(* IEC 61131-3 sources: LASAL/Drive, 5 files *)

(* ---- _DriveAxis1.st ---- *)
FUNCTION GLOBAL TAB DRIVETAB__DRIVEAXIS1
	1$UDINT, TO_UDINT(OFF(L1)-OFF(L0)),L0:
G01:	1$USINT,'U''C''3'' ',
	2$USINT,' '' '' '' ',
	3$USINT,'3''4''V'' ',
	4$USINT,870$DINT,
	5$USINT,3100$DINT,
	6$USINT,12000$DINT,
	7$USINT,2$DINT,
	8$USINT,30$DINT,
	9$USINT,1950$DINT,
	10$USINT,9400$DINT,
	11$USINT,37$DINT,
	12$USINT,6$DINT,
	13$USINT,2$DINT,
	14$USINT,0$DINT,
	15$USINT,330$DINT,
	16$USINT,300$DINT,
	17$USINT,0$DINT,
	18$USINT,0$DINT,
	21$USINT,174$DINT,
	22$USINT,15$DINT,
	23$USINT,35$DINT,
	24$USINT,0$DINT,
	25$USINT,0$DINT,
	26$USINT,0$DINT,
	27$USINT,20$DINT,
G03:	32$USINT,3$DINT,
	33$USINT,50$DINT,
	34$USINT,34$DINT,
	35$USINT,100$DINT,
	36$USINT,200$DINT,
	37$USINT,85$DINT,
	38$USINT,85$DINT,
	39$USINT,0$DINT,
	40$USINT,0$DINT,
	41$USINT,65$DINT,
	42$USINT,235842$DINT,
	43$USINT,2752812$DINT,
	44$USINT,966057170$DINT,
	45$USINT,1111556096$DINT,
	46$USINT,67117569$DINT,
	47$USINT,235842$DINT,
	48$USINT,1$DINT,
	49$USINT,25$DINT,
	168$USINT,60$DINT,
	169$USINT,55$DINT,
	170$USINT,55$DINT,
G04:	50$USINT,4875$DINT,
	51$USINT,1000$DINT,
	52$USINT,50$DINT,
	53$USINT,70$DINT,
	54$USINT,70$DINT,
	55$USINT,40$DINT,
	56$USINT,870$DINT,
	57$USINT,1740$DINT,
	58$USINT,1740$DINT,
G05:	60$USINT,10000$DINT,
	61$USINT,10000$DINT,
	62$USINT,200$DINT,
	63$USINT,1000$DINT,
	64$USINT,80$DINT,
	65$USINT,12000$DINT,
	66$USINT,0$DINT,
G06:	70$USINT,20000$DINT,
	71$USINT,1000$DINT,
	72$USINT,16$DINT,
	73$USINT,1000$DINT,
	74$USINT,0$DINT,
	75$USINT,524288$DINT,
	76$USINT,1$DINT,
G07:	80$USINT,600$DINT,
	81$USINT,0$DINT,
	82$USINT,0$DINT,
	85$USINT,0x00431A06$DINT,
G08:	90$USINT,1000$DINT,
	91$USINT,775$DINT,
	92$USINT,0$DINT,
	93$USINT,3591$DINT,
	94$USINT,0$DINT,
	95$USINT,1000$DINT,
	96$USINT,250$DINT,
	97$USINT,0$DINT,
	98$USINT,0$DINT,
	99$USINT,100$DINT,
	100$USINT,0$DINT,
	101$USINT,100$DINT,
	102$USINT,75$DINT,
	103$USINT,100$DINT,
	104$USINT,0$DINT,
	105$USINT,261$DINT,
	106$USINT,0$DINT,
	107$USINT,0$DINT,
	108$USINT,' '' '' '' ',
	109$USINT,' '' '' '' ',
	110$USINT,' '' '' '' ',
	111$USINT,0$DINT,
	112$USINT,1$DINT,
	113$USINT,0$DINT,
	114$USINT,0$DINT,
	115$USINT,0$DINT,
	116$USINT,0$DINT,
	117$USINT,400$DINT,
	118$USINT,0$DINT,
	119$USINT,2500$DINT,
	120$USINT,20$DINT,
	121$USINT,300$DINT,
	122$USINT,0$DINT,
	173$USINT,0$DINT,L1:
TO_UDINT(OFF(L3)-OFF(L2)),L2:
	01$USINT, OFF(G01),
	03$USINT, OFF(G03),
	04$USINT, OFF(G04),
	05$USINT, OFF(G05),
	06$USINT, OFF(G06),
	07$USINT, OFF(G07),
	08$USINT, OFF(G08),L3:
END_FUNCTION

(* ---- _DriveAxis2.st ---- *)
FUNCTION GLOBAL TAB DRIVETAB__DRIVEAXIS2
	1$UDINT, TO_UDINT(OFF(L1)-OFF(L0)),L0:
G01:	1$USINT,'U''F''6'' ',
	2$USINT,' '' '' '' ',
	3$USINT,'3''4''V'' ',
	4$USINT,2000$DINT,
	5$USINT,4000$DINT,
	6$USINT,7000$DINT,
	7$USINT,2$DINT,
	8$USINT,47$DINT,
	9$USINT,1612$DINT,
	10$USINT,3600$DINT,
	11$USINT,232$DINT,
	13$USINT,2$DINT,
	14$USINT,214$DINT,
	15$USINT,6000$DINT,
	17$USINT,0$DINT,
	18$USINT,0$DINT,
	21$USINT,634$DINT,
	22$USINT,15$DINT,
	23$USINT,35$DINT,
G03:	32$USINT,3$DINT,
	33$USINT,50$DINT,
	35$USINT,20$DINT,
	36$USINT,0$DINT,
	38$USINT,95$DINT,
	41$USINT,65$DINT,
	42$USINT,126550$DINT,
	43$USINT,557767870$DINT,
	44$USINT,33554432$DINT,
	45$USINT,1078001664$DINT,
	46$USINT,67117569$DINT,
	47$USINT,126550$DINT,
	48$USINT,1$DINT,
	49$USINT,15$DINT,
	168$USINT,60$DINT,
	169$USINT,55$DINT,
	170$USINT,65$DINT,
G04:	50$USINT,4030$DINT,
	51$USINT,1000$DINT,
	53$USINT,70$DINT,
	56$USINT,3170$DINT,
	57$USINT,6340$DINT,
	59$USINT,85$DINT,
	167$USINT,100$DINT,
G05:	60$USINT,10000$DINT,
	61$USINT,10000$DINT,
	62$USINT,200$DINT,
	63$USINT,1000$DINT,
	64$USINT,80$DINT,
	65$USINT,2500$DINT,
	66$USINT,0$DINT,
	67$USINT,0$DINT,
	68$USINT,0$DINT,
G06:	70$USINT,20000$DINT,
	71$USINT,1000$DINT,
	72$USINT,16$DINT,
	73$USINT,1000$DINT,
	74$USINT,0$DINT,
	75$USINT,524288$DINT,
	76$USINT,1$DINT,
G08:	90$USINT,1000$DINT,
	91$USINT,775$DINT,
	92$USINT,0$DINT,
	93$USINT,2567$DINT,
	94$USINT,0$DINT,
	95$USINT,1000$DINT,
	99$USINT,80$DINT,
	103$USINT,1$DINT,
	105$USINT,951$DINT,
	108$USINT,' '' '' '' ',
	109$USINT,' '' '' '' ',
	110$USINT,' '' '' '' ',
	114$USINT,0$DINT,
	115$USINT,0$DINT,
	116$USINT,0$DINT,
	117$USINT,400$DINT,
	118$USINT,0$DINT,
	119$USINT,2500$DINT,
	120$USINT,20$DINT,
	121$USINT,300$DINT,
	124$USINT,1163207552$DINT,
	164$USINT,0$DINT,
	165$USINT,0$DINT,
	173$USINT,12$DINT,
G14:	127$USINT,0$DINT,
	128$USINT,100$DINT,
	129$USINT,100$DINT,
	130$USINT,100$DINT,
	131$USINT,100$DINT,
	132$USINT,100$DINT,
	133$USINT,100$DINT,
	134$USINT,100$DINT,
	135$USINT,100$DINT,
	136$USINT,100$DINT,
	137$USINT,100$DINT,
	138$USINT,100$DINT,
	139$USINT,100$DINT,
	140$USINT,100$DINT,
	141$USINT,100$DINT,
	142$USINT,100$DINT,
	143$USINT,100$DINT,
	144$USINT,100$DINT,
	145$USINT,100$DINT,
	146$USINT,100$DINT,
	147$USINT,100$DINT,
	148$USINT,100$DINT,
	149$USINT,100$DINT,
	150$USINT,100$DINT,
	151$USINT,100$DINT,
	152$USINT,100$DINT,
	153$USINT,100$DINT,
	154$USINT,100$DINT,
	155$USINT,100$DINT,
	156$USINT,100$DINT,
	157$USINT,100$DINT,
	158$USINT,100$DINT,
	159$USINT,100$DINT,L1:
TO_UDINT(OFF(L3)-OFF(L2)),L2:
	01$USINT, OFF(G01),
	03$USINT, OFF(G03),
	04$USINT, OFF(G04),
	05$USINT, OFF(G05),
	06$USINT, OFF(G06),
	08$USINT, OFF(G08),
	14$USINT, OFF(G14),L3:
END_FUNCTION

(* ---- _DriveAxis3.st ---- *)
FUNCTION GLOBAL TAB DRIVETAB__DRIVEAXIS3
	1$UDINT, TO_UDINT(OFF(L1)-OFF(L0)),L0:
G01:	1$USINT,'U''M''3''S',
	2$USINT,' '' '' '' ',
	3$USINT,'3''4''V'' ',
	4$USINT,1500$DINT,
	5$USINT,5000$DINT,
	6$USINT,2000$DINT,
	7$USINT,2$DINT,
	8$USINT,95$DINT,
	9$USINT,4680$DINT,
	10$USINT,11000$DINT,
	11$USINT,589$DINT,
	12$USINT,6$DINT,
	13$USINT,2$DINT,
	14$USINT,115$DINT,
	15$USINT,6000$DINT,
	16$USINT,300$DINT,
	17$USINT,0$DINT,
	18$USINT,0$DINT,
	21$USINT,300$DINT,
	22$USINT,15$DINT,
	23$USINT,35$DINT,
	24$USINT,0$DINT,
	25$USINT,0$DINT,
	26$USINT,0$DINT,
	27$USINT,20$DINT,
G03:	32$USINT,3$DINT,
	33$USINT,50$DINT,
	34$USINT,34$DINT,
	35$USINT,100$DINT,
	36$USINT,200$DINT,
	37$USINT,85$DINT,
	38$USINT,85$DINT,
	39$USINT,0$DINT,
	40$USINT,0$DINT,
	41$USINT,65$DINT,
	42$USINT,71519$DINT,
	43$USINT,2752812$DINT,
	44$USINT,966057170$DINT,
	45$USINT,1111556096$DINT,
	46$USINT,67117569$DINT,
	47$USINT,71519$DINT,
	48$USINT,1$DINT,
	49$USINT,25$DINT,
	168$USINT,60$DINT,
	169$USINT,55$DINT,
	170$USINT,55$DINT,
G04:	50$USINT,11700$DINT,
	51$USINT,1000$DINT,
	52$USINT,50$DINT,
	53$USINT,70$DINT,
	54$USINT,70$DINT,
	55$USINT,40$DINT,
	56$USINT,1500$DINT,
	57$USINT,3000$DINT,
	58$USINT,3000$DINT,
G05:	60$USINT,10000$DINT,
	61$USINT,10000$DINT,
	62$USINT,200$DINT,
	63$USINT,1000$DINT,
	64$USINT,80$DINT,
	65$USINT,2000$DINT,
	66$USINT,0$DINT,
G06:	70$USINT,20000$DINT,
	71$USINT,1000$DINT,
	72$USINT,16$DINT,
	73$USINT,1000$DINT,
	74$USINT,0$DINT,
	75$USINT,524288$DINT,
	76$USINT,1$DINT,
G07:	80$USINT,600$DINT,
	81$USINT,0$DINT,
	82$USINT,0$DINT,
G08:	90$USINT,1000$DINT,
	91$USINT,775$DINT,
	92$USINT,0$DINT,
	93$USINT,3591$DINT,
	94$USINT,0$DINT,
	95$USINT,1000$DINT,
	96$USINT,250$DINT,
	97$USINT,0$DINT,
	98$USINT,0$DINT,
	99$USINT,100$DINT,
	100$USINT,0$DINT,
	101$USINT,100$DINT,
	102$USINT,75$DINT,
	103$USINT,100$DINT,
	104$USINT,0$DINT,
	105$USINT,450$DINT,
	106$USINT,0$DINT,
	107$USINT,0$DINT,
	108$USINT,' '' '' '' ',
	109$USINT,' '' '' '' ',
	110$USINT,' '' '' '' ',
	111$USINT,0$DINT,
	112$USINT,1$DINT,
	113$USINT,0$DINT,
	114$USINT,0$DINT,
	115$USINT,0$DINT,
	116$USINT,0$DINT,
	117$USINT,400$DINT,
	118$USINT,0$DINT,
	119$USINT,2500$DINT,
	120$USINT,20$DINT,
	121$USINT,300$DINT,
	122$USINT,0$DINT,
	173$USINT,0$DINT,L1:
TO_UDINT(OFF(L3)-OFF(L2)),L2:
	01$USINT, OFF(G01),
	03$USINT, OFF(G03),
	04$USINT, OFF(G04),
	05$USINT, OFF(G05),
	06$USINT, OFF(G06),
	07$USINT, OFF(G07),
	08$USINT, OFF(G08),L3:
END_FUNCTION

(* ---- _DriveAxis4.st ---- *)
FUNCTION GLOBAL TAB DRIVETAB__DRIVEAXIS4
	1$UDINT, TO_UDINT(OFF(L1)-OFF(L0)),L0:
G01:	1$USINT,'U''M''3''S',
	2$USINT,' '' '' '' ',
	3$USINT,'3''4''V'' ',
	4$USINT,1500$DINT,
	5$USINT,5000$DINT,
	6$USINT,1000$DINT,
	7$USINT,2$DINT,
	8$USINT,95$DINT,
	9$USINT,4680$DINT,
	10$USINT,11000$DINT,
	11$USINT,589$DINT,
	13$USINT,2$DINT,
	14$USINT,337$DINT,
	15$USINT,6000$DINT,
	17$USINT,0$DINT,
	18$USINT,0$DINT,
	21$USINT,300$DINT,
	22$USINT,15$DINT,
	23$USINT,35$DINT,
G03:	32$USINT,3$DINT,
	33$USINT,50$DINT,
	35$USINT,15$DINT,
	36$USINT,200$DINT,
	38$USINT,95$DINT,
	41$USINT,65$DINT,
	42$USINT,71519$DINT,
	43$USINT,2752812$DINT,
	44$USINT,0$DINT,
	45$USINT,1111556096$DINT,
	46$USINT,67117569$DINT,
	47$USINT,71519$DINT,
	48$USINT,1$DINT,
	49$USINT,25$DINT,
	168$USINT,55$DINT,
	169$USINT,52$DINT,
	170$USINT,65$DINT,
G04:	50$USINT,11700$DINT,
	51$USINT,1000$DINT,
	53$USINT,70$DINT,
	56$USINT,1500$DINT,
	57$USINT,3000$DINT,
	59$USINT,85$DINT,
	167$USINT,100$DINT,
G05:	60$USINT,5000$DINT,
	61$USINT,10000$DINT,
	62$USINT,200$DINT,
	63$USINT,1000$DINT,
	64$USINT,80$DINT,
	65$USINT,1000$DINT,
	66$USINT,0$DINT,
	67$USINT,0$DINT,
	68$USINT,0$DINT,
G06:	70$USINT,10000$DINT,
	71$USINT,1000$DINT,
	72$USINT,16$DINT,
	73$USINT,1000$DINT,
	74$USINT,0$DINT,
	75$USINT,524288$DINT,
	76$USINT,1$DINT,
G08:	90$USINT,1000$DINT,
	91$USINT,775$DINT,
	92$USINT,0$DINT,
	93$USINT,2567$DINT,
	94$USINT,0$DINT,
	95$USINT,1000$DINT,
	99$USINT,100$DINT,
	103$USINT,100$DINT,
	105$USINT,650$DINT,
	108$USINT,' '' '' '' ',
	109$USINT,' '' '' '' ',
	110$USINT,' '' '' '' ',
	114$USINT,0$DINT,
	115$USINT,0$DINT,
	116$USINT,0$DINT,
	117$USINT,400$DINT,
	118$USINT,0$DINT,
	119$USINT,2500$DINT,
	120$USINT,20$DINT,
	121$USINT,300$DINT,
	124$USINT,1217332736$DINT,
	164$USINT,0$DINT,
	165$USINT,0$DINT,
	173$USINT,0$DINT,
G14:	127$USINT,0$DINT,
	128$USINT,100$DINT,
	129$USINT,100$DINT,
	130$USINT,100$DINT,
	131$USINT,100$DINT,
	132$USINT,100$DINT,
	133$USINT,100$DINT,
	134$USINT,100$DINT,
	135$USINT,100$DINT,
	136$USINT,100$DINT,
	137$USINT,100$DINT,
	138$USINT,100$DINT,
	139$USINT,100$DINT,
	140$USINT,100$DINT,
	141$USINT,100$DINT,
	142$USINT,100$DINT,
	143$USINT,100$DINT,
	144$USINT,100$DINT,
	145$USINT,100$DINT,
	146$USINT,100$DINT,
	147$USINT,100$DINT,
	148$USINT,100$DINT,
	149$USINT,100$DINT,
	150$USINT,100$DINT,
	151$USINT,100$DINT,
	152$USINT,100$DINT,
	153$USINT,100$DINT,
	154$USINT,100$DINT,
	155$USINT,100$DINT,
	156$USINT,100$DINT,
	157$USINT,100$DINT,
	158$USINT,100$DINT,
	159$USINT,100$DINT,L1:
TO_UDINT(OFF(L3)-OFF(L2)),L2:
	01$USINT, OFF(G01),
	03$USINT, OFF(G03),
	04$USINT, OFF(G04),
	05$USINT, OFF(G05),
	06$USINT, OFF(G06),
	08$USINT, OFF(G08),
	14$USINT, OFF(G14),L3:
END_FUNCTION

(* ---- DRIVETAB03.st ---- *)
FUNCTION GLOBAL TAB DRIVETAB3
	1$UDINT, TO_UDINT(OFF(L1)-OFF(L0)),L0:
G01:	1$USINT,'U''C''3'' ',
	2$USINT,' '' '' '' ',
	3$USINT,'3''4''V'' ',
	4$USINT,870$DINT,
	5$USINT,3100$DINT,
	6$USINT,12000$DINT,
	7$USINT,2$DINT,
	8$USINT,30$DINT,
	9$USINT,1950$DINT,
	10$USINT,9400$DINT,
	11$USINT,37$DINT,
	13$USINT,2$DINT,
	14$USINT,288$DINT,
	15$USINT,330$DINT,
	17$USINT,0$DINT,
	18$USINT,0$DINT,
	21$USINT,174$DINT,
	22$USINT,15$DINT,
	23$USINT,35$DINT,
G03:	32$USINT,-2$DINT,
	33$USINT,50$DINT,
	35$USINT,20$DINT,
	36$USINT,0$DINT,
	38$USINT,85$DINT,
	41$USINT,65$DINT,
	42$USINT,10000$DINT,
	43$USINT,2752812$DINT,
	44$USINT,0$DINT,
	45$USINT,1111556096$DINT,
	46$USINT,67117569$DINT,
	47$USINT,235842$DINT,
	48$USINT,1$DINT,
	49$USINT,0$DINT,
	168$USINT,55$DINT,
	169$USINT,52$DINT,
	170$USINT,65$DINT,
G04:	50$USINT,4875$DINT,
	51$USINT,1000$DINT,
	53$USINT,70$DINT,
	56$USINT,870$DINT,
	57$USINT,3000$DINT,
	59$USINT,85$DINT,
	167$USINT,100$DINT,
G05:	60$USINT,9000$DINT,
	61$USINT,0$DINT,
	62$USINT,200$DINT,
	63$USINT,1000$DINT,
	64$USINT,80$DINT,
	65$USINT,12000$DINT,
	66$USINT,0$DINT,
	67$USINT,0$DINT,
	68$USINT,0$DINT,
G06:	70$USINT,20000$DINT,
	71$USINT,1000$DINT,
	72$USINT,16$DINT,
	73$USINT,1000$DINT,
	74$USINT,0$DINT,
	75$USINT,524288$DINT,
	76$USINT,1$DINT,
G08:	90$USINT,1000$DINT,
	91$USINT,517$DINT,
	92$USINT,0$DINT,
	93$USINT,2567$DINT,
	94$USINT,0$DINT,
	95$USINT,1000$DINT,
	99$USINT,100$DINT,
	103$USINT,100$DINT,
	105$USINT,500$DINT,
	108$USINT,' '' '' '' ',
	109$USINT,' '' '' '' ',
	110$USINT,' '' '' '' ',
	114$USINT,0$DINT,
	115$USINT,0$DINT,
	116$USINT,0$DINT,
	117$USINT,400$DINT,
	118$USINT,0$DINT,
	119$USINT,2500$DINT,
	120$USINT,20$DINT,
	121$USINT,300$DINT,
	124$USINT,1217334272$DINT,
	164$USINT,0$DINT,
	165$USINT,0$DINT,
	173$USINT,0$DINT,
G14:	127$USINT,0$DINT,
	128$USINT,100$DINT,
	129$USINT,100$DINT,
	130$USINT,100$DINT,
	131$USINT,100$DINT,
	132$USINT,100$DINT,
	133$USINT,100$DINT,
	134$USINT,100$DINT,
	135$USINT,100$DINT,
	136$USINT,100$DINT,
	137$USINT,100$DINT,
	138$USINT,100$DINT,
	139$USINT,100$DINT,
	140$USINT,100$DINT,
	141$USINT,100$DINT,
	142$USINT,100$DINT,
	143$USINT,100$DINT,
	144$USINT,100$DINT,
	145$USINT,100$DINT,
	146$USINT,100$DINT,
	147$USINT,100$DINT,
	148$USINT,100$DINT,
	149$USINT,100$DINT,
	150$USINT,100$DINT,
	151$USINT,100$DINT,
	152$USINT,100$DINT,
	153$USINT,100$DINT,
	154$USINT,100$DINT,
	155$USINT,100$DINT,
	156$USINT,100$DINT,
	157$USINT,100$DINT,
	158$USINT,100$DINT,
	159$USINT,100$DINT,L1:
TO_UDINT(OFF(L3)-OFF(L2)),L2:
	01$USINT, OFF(G01),
	03$USINT, OFF(G03),
	04$USINT, OFF(G04),
	05$USINT, OFF(G05),
	06$USINT, OFF(G06),
	08$USINT, OFF(G08),
	14$USINT, OFF(G14),L3:
END_FUNCTION
